(* IEC 61131-3 sources: codesys-to-astra/src/DUTs, 5 files *)

(* ---- E_C2aDecimalSeparator.dut.st ---- *)
// Назначение: разделитель целой и дробной части для F_C2aRealToStringFormat — аналог
//             перечисления DECIMAL_SEPARATOR OwenStringUtils (DOT = 0, COMMA = 1, USINT; документ ОВЕН v3.0,
//             табл. 3.2.2, с. 9).
// Автор:      kr0nsch
// Версия:     0.1.0
// Документ:   docs/LIBMAP.md
{attribute 'qualified_only'}
{attribute 'strict'}
TYPE E_C2aDecimalSeparator :
(
    DOT := 0,       // точка
    COMMA := 1      // запятая
) USINT;
END_TYPE

(* ---- E_C2aMx210Status.dut.st ---- *)
// Назначение: состояние измерения МВ210-101 по коду ошибки в регистре значения (РЭ МВ210-101 v1.41,
//             табл. 6.9, с. 36). Положение кода в регистрах FLOAT32/INT16 по РЭ однозначно не следует — сверить
//             на модуле (docs/HARDWARE_VALIDATION.md).
// Автор:      kr0nsch
// Версия:     0.1.0
// Документ:   docs/IO.md
{attribute 'qualified_only'}
TYPE E_C2aMx210Status :
(
    Ok := 0,                // передаётся результат измерения
    Invalid := 16#F0,       // значение заведомо неверно
    NotReady := 16#F6,      // данные не готовы
    SensorOff := 16#F7,     // датчик отключён
    ColdJunctionHigh := 16#F8,  // велика температура свободных концов ТП
    ColdJunctionLow := 16#F9,   // мала температура свободных концов ТП
    TooHigh := 16#FA,       // значение слишком велико
    TooLow := 16#FB,        // значение слишком мало
    ShortCircuit := 16#FC,  // короткое замыкание датчика
    SensorBreak := 16#FD,   // обрыв датчика
    AdcFailure := 16#FE,    // нет связи с АЦП
    BadCalibration := 16#FF // некорректный калибровочный коэффициент
) BYTE;
END_TYPE

(* ---- E_C2aWordOrder.dut.st ---- *)
// Назначение: порядок слов 32-битного значения в двух регистрах Modbus (канал REGUL отдаёт
//             ARRAY OF WORD, DPA-302.1 с. 15–16). Порядок слов FLOAT32 Mx210 через драйвер REGUL не сверен —
//             docs/HARDWARE_VALIDATION.md.
// Автор:      kr0nsch
// Версия:     0.1.0
// Документ:   docs/IO.md
{attribute 'qualified_only'}
TYPE E_C2aWordOrder :
(
    HighWordFirst := 0,     // старшее слово в первом регистре
    LowWordFirst := 1       // младшее слово в первом регистре
) USINT;
END_TYPE

(* ---- ST_C2aDateTime.dut.st ---- *)
// Назначение: дата и время по каналам узла OwenRTC (Targets v3.4, табл. 4.1, с. 10–11).
// Автор:      kr0nsch
// Версия:     0.1.0
// Документ:   docs/LIBMAP.md
TYPE ST_C2aDateTime :
STRUCT
    uiYear : UINT;          // год
    usiMonth : USINT;       // месяц 1..12
    usiDay : USINT;         // день 1..31
    usiHour : USINT;        // час 0..23
    usiMinute : USINT;      // минута 0..59
    usiSecond : USINT;      // секунда 0..59
    usiDayOfWeek : USINT;   // день недели: 1 — понедельник, 7 — воскресенье
END_STRUCT
END_TYPE

(* ---- U_C2aReal32.dut.st ---- *)
// Назначение: 32 бита как REAL или DWORD — распаковка FLOAT32 из двух регистров Modbus.
// Автор:      kr0nsch
// Версия:     0.1.0
// Документ:   docs/IO.md
TYPE U_C2aReal32 :
UNION
    rValue : REAL;      // значение с плавающей точкой
    dwValue : DWORD;    // то же как 32 бита
END_UNION
END_TYPE
